Fanuc KAREL source: KT00725.KL

PROGRAM KT00725
%NOLOCKGROUP
VAR
  P1: JOINTPOS
  P2: JOINTPOS
  OUT: INTEGER
BEGIN
  OUT = ARRAY_LEN(P1)
END KT00725
